(* IEC 61131-3 sources: trust-platform/examples/tutorials/10_unit_testing_101/sources, 2 files *)

(* ---- main.st ---- *)
FUNCTION LIMIT_ADD : INT
VAR_INPUT
    A : INT;
    B : INT;
    MAX_VALUE : INT;
END_VAR
VAR
    SUM : INT;
END_VAR

SUM := A + B;
IF SUM > MAX_VALUE THEN
    LIMIT_ADD := MAX_VALUE;
ELSE
    LIMIT_ADD := SUM;
END_IF;
END_FUNCTION

FUNCTION SCALE_RAW_TO_PERCENT : REAL
VAR_INPUT
    RAW : INT;
END_VAR

SCALE_RAW_TO_PERCENT := INT_TO_REAL(IN := RAW) * REAL#0.1;
END_FUNCTION

FUNCTION_BLOCK FB_START_STOP
VAR_INPUT
    StartCmd : BOOL;
    StopCmd : BOOL;
END_VAR
VAR_OUTPUT
    Running : BOOL;
END_VAR

IF StopCmd THEN
    Running := FALSE;
ELSIF StartCmd THEN
    Running := TRUE;
END_IF;
END_FUNCTION_BLOCK

(* ---- tests.st ---- *)
TEST_PROGRAM TEST_LIMIT_ADD_AND_SCALING
ASSERT_EQUAL(
    EXPECTED := INT#7,
    ACTUAL := LIMIT_ADD(A := INT#3, B := INT#4, MAX_VALUE := INT#10)
);
ASSERT_EQUAL(
    EXPECTED := INT#5,
    ACTUAL := LIMIT_ADD(A := INT#3, B := INT#4, MAX_VALUE := INT#5)
);
ASSERT_EQUAL(
    EXPECTED := INT#-2,
    ACTUAL := LIMIT_ADD(A := INT#-3, B := INT#1, MAX_VALUE := INT#100)
);
(* REAL assertions should use tolerance for stable behavior. *)
ASSERT_NEAR(
    EXPECTED := REAL#37.5,
    ACTUAL := SCALE_RAW_TO_PERCENT(RAW := INT#375),
    DELTA := REAL#0.01
);
ASSERT_TRUE(IN := LIMIT_ADD(A := INT#2, B := INT#2, MAX_VALUE := INT#5) = INT#4);
ASSERT_FALSE(IN := LIMIT_ADD(A := INT#2, B := INT#2, MAX_VALUE := INT#3) = INT#4);
END_TEST_PROGRAM

TEST_FUNCTION_BLOCK TEST_FB_START_STOP_SEQUENCE
VAR
    DUT : FB_START_STOP;
END_VAR

(* Cycle 1: idle state, output should stay FALSE. *)
DUT(StartCmd := FALSE, StopCmd := FALSE);
ASSERT_FALSE(DUT.Running);

(* Cycle 2: start command latches Running TRUE. *)
DUT(StartCmd := TRUE, StopCmd := FALSE);
ASSERT_TRUE(DUT.Running);

(* Cycle 3: no input change keeps the latched state. *)
DUT(StartCmd := FALSE, StopCmd := FALSE);
ASSERT_TRUE(DUT.Running);

(* Cycle 4: stop command resets Running to FALSE. *)
DUT(StartCmd := FALSE, StopCmd := TRUE);
ASSERT_FALSE(DUT.Running);
END_TEST_FUNCTION_BLOCK
